(* Cycle Allowed only if both safety conditions are True *)

PROGRAM main
  VAR
    InputA AT %IX0.2 : BOOL;
    InputB AT %IX0.3 : BOOL; (* Guard Closed *)
    Output AT %MX0.0 : BOOL;
  END_VAR

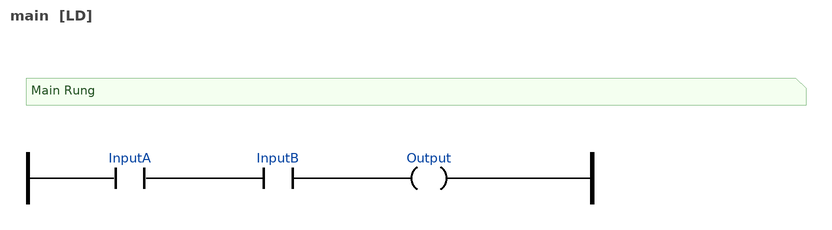
(* LD diagram, written out as Structured Text *)
(* Main Rung *)
Output := InputA AND InputB;
END_PROGRAM
